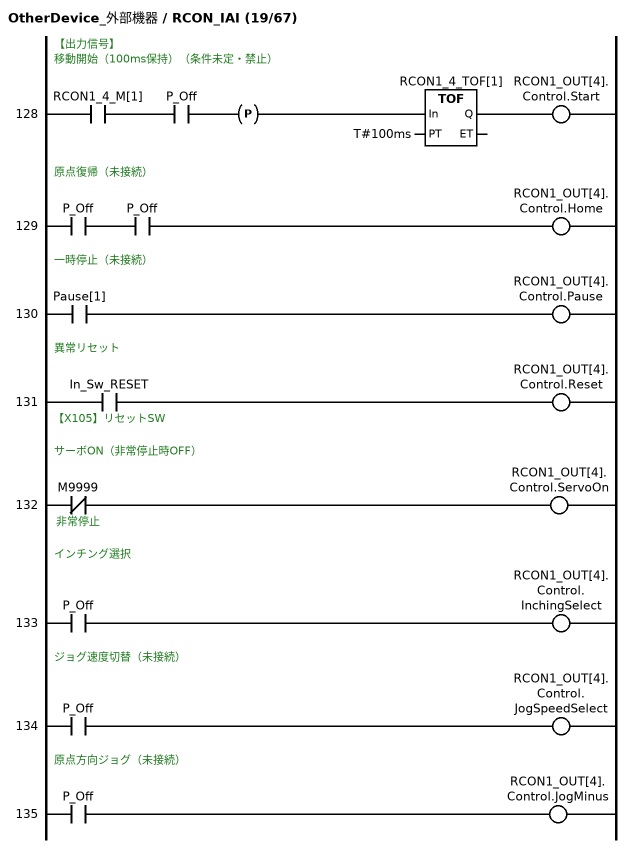
(* [picture p96: OtherDevice_外部機器 / RCON_IAI, rungs 128-135] *)
(* Rung 128: 【出力信号】 / 移動開始（100ms保持）（条件未定・禁止） *)
_e13(CLK := RCON1_4_M[1] AND P_Off);
RCON1_4_TOF[1](In := _e13.Q, PT := T#100ms);
RCON1_OUT[4].Control.Start := RCON1_4_TOF[1].Q;
(* Rung 129: 原点復帰（未接続） *)
RCON1_OUT[4].Control.Home := P_Off AND P_Off;
(* Rung 130: 一時停止（未接続） *)
RCON1_OUT[4].Control.Pause := Pause[1];
(* Rung 131: 異常リセット *)
RCON1_OUT[4].Control.Reset := In_Sw_RESET;
(* Rung 132: サーボON（非常停止時OFF） *)
RCON1_OUT[4].Control.ServoOn := NOT M9999;
(* Rung 133: インチング選択 *)
RCON1_OUT[4].Control.InchingSelect := P_Off;
(* Rung 134: ジョグ速度切替（未接続） *)
RCON1_OUT[4].Control.JogSpeedSelect := P_Off;
(* Rung 135: 原点方向ジョグ（未接続） *)
RCON1_OUT[4].Control.JogMinus := P_Off;

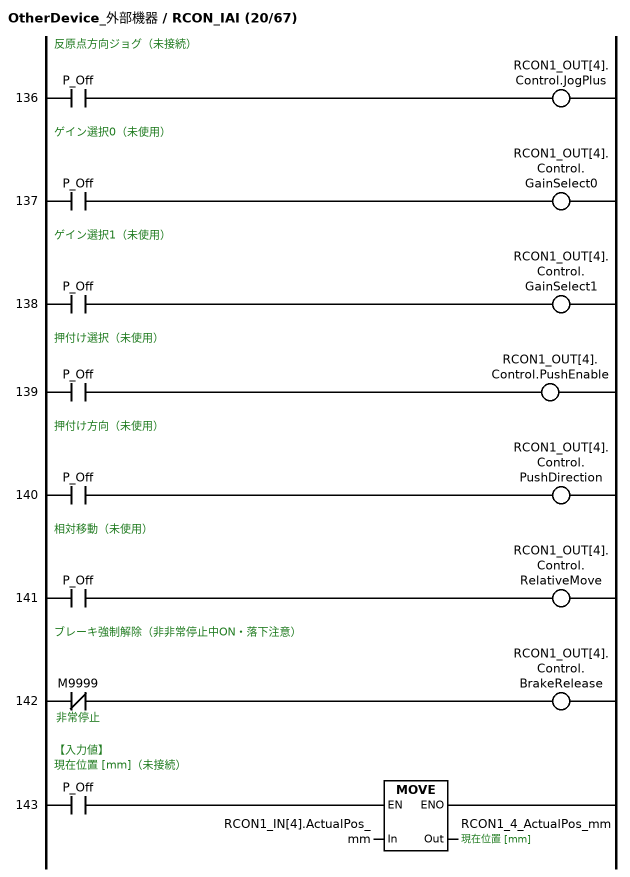
(* Rung 136: 反原点方向ジョグ（未接続） *)
RCON1_OUT[4].Control.JogPlus := P_Off;
(* Rung 137: ゲイン選択0（未使用） *)
RCON1_OUT[4].Control.GainSelect0 := P_Off;
(* Rung 138: ゲイン選択1（未使用） *)
RCON1_OUT[4].Control.GainSelect1 := P_Off;
(* Rung 139: 押付け選択（未使用） *)
RCON1_OUT[4].Control.PushEnable := P_Off;
(* Rung 140: 押付け方向（未使用） *)
RCON1_OUT[4].Control.PushDirection := P_Off;
(* Rung 141: 相対移動（未使用） *)
RCON1_OUT[4].Control.RelativeMove := P_Off;
(* Rung 142: ブレーキ強制解除（非非常停止中ON・落下注意） *)
RCON1_OUT[4].Control.BrakeRelease := NOT M9999;
(* Rung 143: 【入力値】 / 現在位置 [mm]（未接続） *)
IF P_Off THEN RCON1_4_ActualPos_mm := RCON1_IN[4].ActualPos_mm; END_IF;

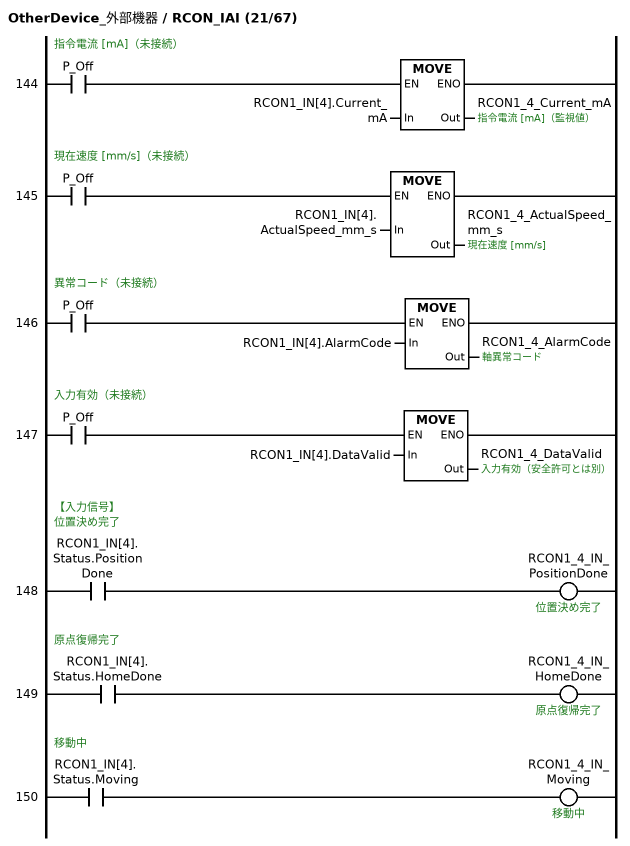
(* Rung 144: 指令電流 [mA]（未接続） *)
IF P_Off THEN RCON1_4_Current_mA := RCON1_IN[4].Current_mA; END_IF;
(* Rung 145: 現在速度 [mm/s]（未接続） *)
IF P_Off THEN RCON1_4_ActualSpeed_mm_s := RCON1_IN[4].ActualSpeed_mm_s; END_IF;
(* Rung 146: 異常コード（未接続） *)
IF P_Off THEN RCON1_4_AlarmCode := RCON1_IN[4].AlarmCode; END_IF;
(* Rung 147: 入力有効（未接続） *)
IF P_Off THEN RCON1_4_DataValid := RCON1_IN[4].DataValid; END_IF;
(* Rung 148: 【入力信号】 / 位置決め完了 *)
RCON1_4_IN_PositionDone := RCON1_IN[4].Status.PositionDone;
(* Rung 149: 原点復帰完了 *)
RCON1_4_IN_HomeDone := RCON1_IN[4].Status.HomeDone;
(* Rung 150: 移動中 *)
RCON1_4_IN_Moving := RCON1_IN[4].Status.Moving;

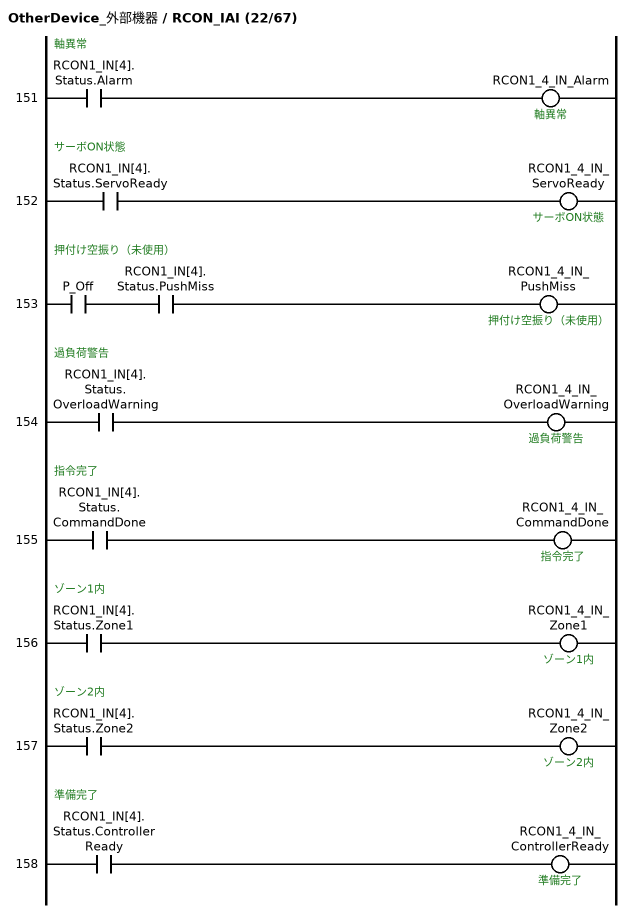
(* Rung 151: 軸異常 *)
RCON1_4_IN_Alarm := RCON1_IN[4].Status.Alarm;
(* Rung 152: サーボON状態 *)
RCON1_4_IN_ServoReady := RCON1_IN[4].Status.ServoReady;
(* Rung 153: 押付け空振り（未使用） *)
RCON1_4_IN_PushMiss := P_Off AND RCON1_IN[4].Status.PushMiss;
(* Rung 154: 過負荷警告 *)
RCON1_4_IN_OverloadWarning := RCON1_IN[4].Status.OverloadWarning;
(* Rung 155: 指令完了 *)
RCON1_4_IN_CommandDone := RCON1_IN[4].Status.CommandDone;
(* Rung 156: ゾーン1内 *)
RCON1_4_IN_Zone1 := RCON1_IN[4].Status.Zone1;
(* Rung 157: ゾーン2内 *)
RCON1_4_IN_Zone2 := RCON1_IN[4].Status.Zone2;
(* Rung 158: 準備完了 *)
RCON1_4_IN_ControllerReady := RCON1_IN[4].Status.ControllerReady;

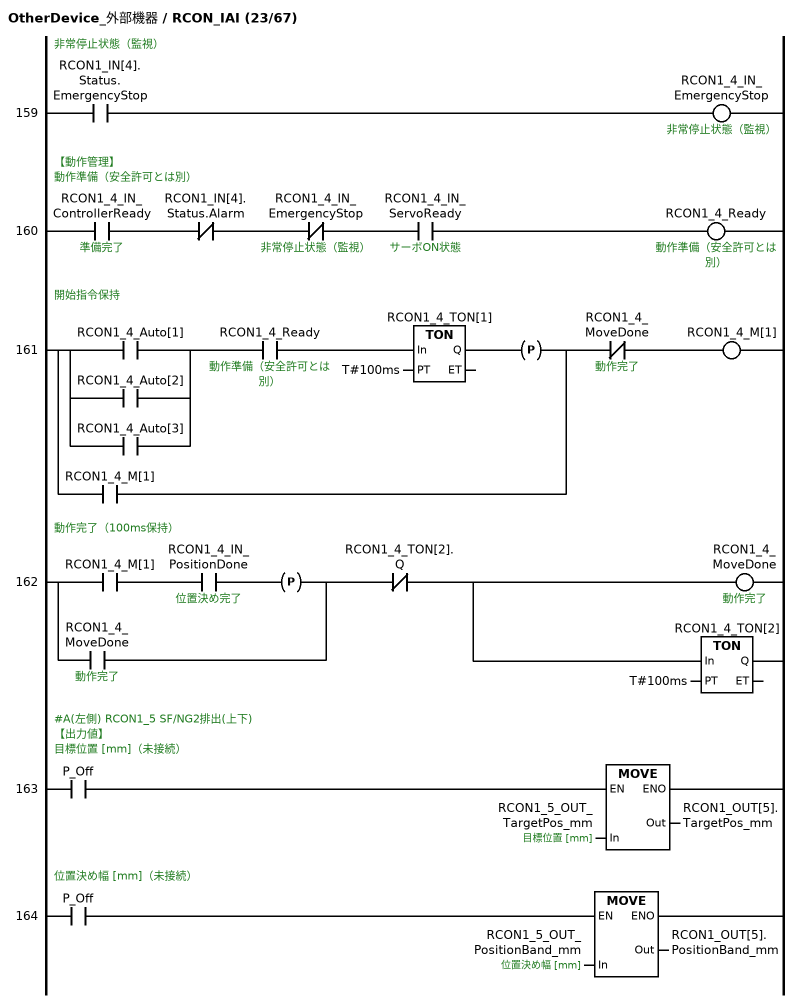
(* Rung 159: 非常停止状態（監視） *)
RCON1_4_IN_EmergencyStop := RCON1_IN[4].Status.EmergencyStop;
(* Rung 160: 【動作管理】 / 動作準備（安全許可とは別） *)
RCON1_4_Ready := RCON1_4_IN_ControllerReady AND NOT RCON1_IN[4].Status.Alarm AND NOT RCON1_4_IN_EmergencyStop AND RCON1_4_IN_ServoReady;
(* Rung 161: 開始指令保持 *)
RCON1_4_TON[1](In := (RCON1_4_Auto[1] OR RCON1_4_Auto[2] OR RCON1_4_Auto[3]) AND RCON1_4_Ready, PT := T#100ms);
_e14(CLK := RCON1_4_TON[1].Q);
RCON1_4_M[1] := (_e14.Q OR RCON1_4_M[1]) AND NOT RCON1_4_MoveDone;
(* Rung 162: 動作完了（100ms保持） *)
_e15(CLK := RCON1_4_M[1] AND RCON1_4_IN_PositionDone);
_p16 := (_e15.Q OR RCON1_4_MoveDone) AND NOT RCON1_4_TON[2].Q;
RCON1_4_MoveDone := _p16;
RCON1_4_TON[2](In := _p16, PT := T#100ms);
(* Rung 163: #A(左側) RCON1_5 SF/NG2排出(上下) / 【出力値】 / 目標位置 [mm]（未接続） *)
IF P_Off THEN RCON1_OUT[5].TargetPos_mm := RCON1_5_OUT_TargetPos_mm; END_IF;
(* Rung 164: 位置決め幅 [mm]（未接続） *)
IF P_Off THEN RCON1_OUT[5].PositionBand_mm := RCON1_5_OUT_PositionBand_mm; END_IF;

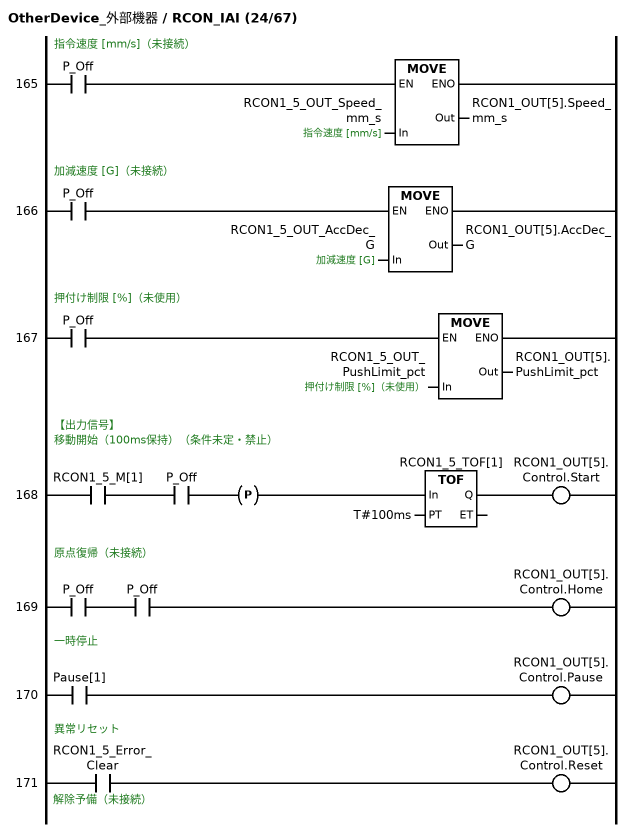
(* Rung 165: 指令速度 [mm/s]（未接続） *)
IF P_Off THEN RCON1_OUT[5].Speed_mm_s := RCON1_5_OUT_Speed_mm_s; END_IF;
(* Rung 166: 加減速度 [G]（未接続） *)
IF P_Off THEN RCON1_OUT[5].AccDec_G := RCON1_5_OUT_AccDec_G; END_IF;
(* Rung 167: 押付け制限 [%]（未使用） *)
IF P_Off THEN RCON1_OUT[5].PushLimit_pct := RCON1_5_OUT_PushLimit_pct; END_IF;
(* Rung 168: 【出力信号】 / 移動開始（100ms保持）（条件未定・禁止） *)
_e17(CLK := RCON1_5_M[1] AND P_Off);
RCON1_5_TOF[1](In := _e17.Q, PT := T#100ms);
RCON1_OUT[5].Control.Start := RCON1_5_TOF[1].Q;
(* Rung 169: 原点復帰（未接続） *)
RCON1_OUT[5].Control.Home := P_Off AND P_Off;
(* Rung 170: 一時停止 *)
RCON1_OUT[5].Control.Pause := Pause[1];
(* Rung 171: 異常リセット *)
RCON1_OUT[5].Control.Reset := RCON1_5_Error_Clear;

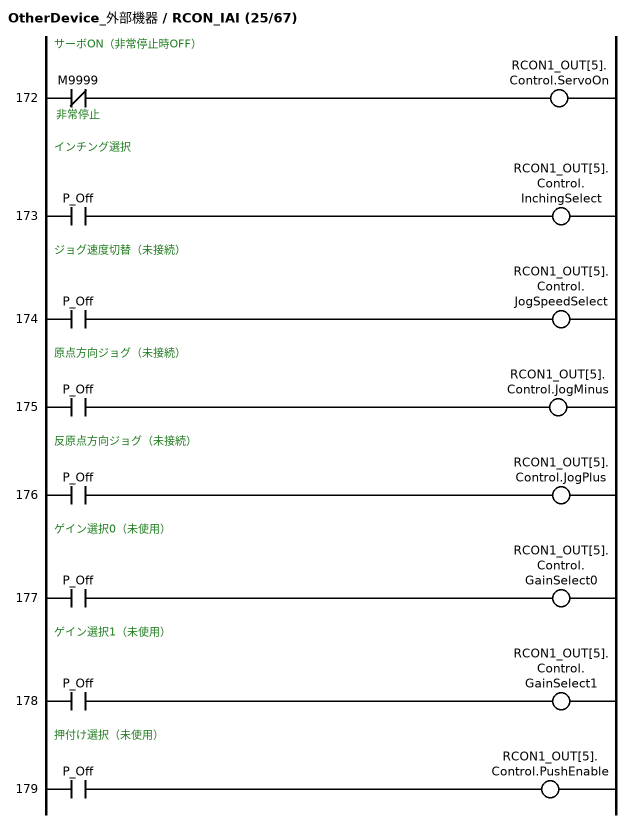
(* Rung 172: サーボON（非常停止時OFF） *)
RCON1_OUT[5].Control.ServoOn := NOT M9999;
(* Rung 173: インチング選択 *)
RCON1_OUT[5].Control.InchingSelect := P_Off;
(* Rung 174: ジョグ速度切替（未接続） *)
RCON1_OUT[5].Control.JogSpeedSelect := P_Off;
(* Rung 175: 原点方向ジョグ（未接続） *)
RCON1_OUT[5].Control.JogMinus := P_Off;
(* Rung 176: 反原点方向ジョグ（未接続） *)
RCON1_OUT[5].Control.JogPlus := P_Off;
(* Rung 177: ゲイン選択0（未使用） *)
RCON1_OUT[5].Control.GainSelect0 := P_Off;
(* Rung 178: ゲイン選択1（未使用） *)
RCON1_OUT[5].Control.GainSelect1 := P_Off;
(* Rung 179: 押付け選択（未使用） *)
RCON1_OUT[5].Control.PushEnable := P_Off;

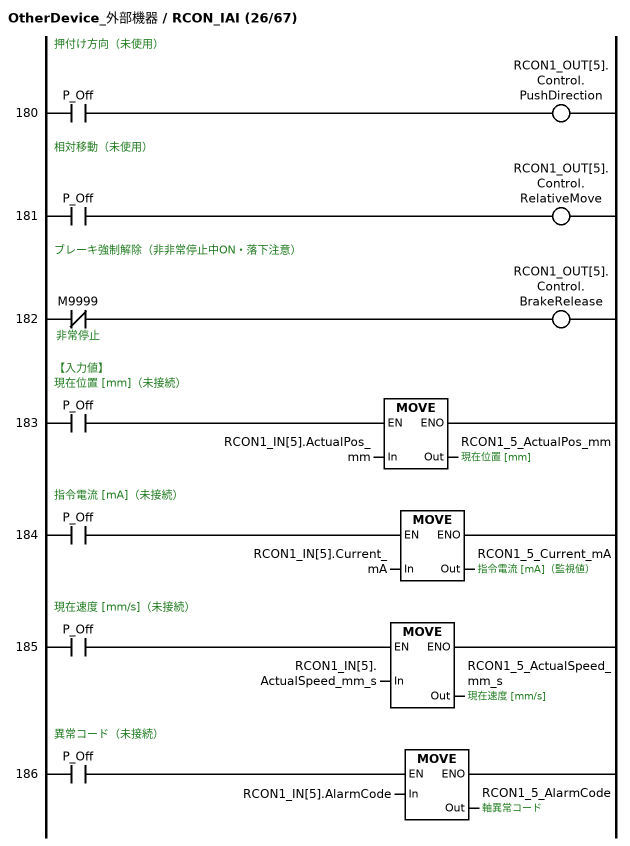
(* Rung 180: 押付け方向（未使用） *)
RCON1_OUT[5].Control.PushDirection := P_Off;
(* Rung 181: 相対移動（未使用） *)
RCON1_OUT[5].Control.RelativeMove := P_Off;
(* Rung 182: ブレーキ強制解除（非非常停止中ON・落下注意） *)
RCON1_OUT[5].Control.BrakeRelease := NOT M9999;
(* Rung 183: 【入力値】 / 現在位置 [mm]（未接続） *)
IF P_Off THEN RCON1_5_ActualPos_mm := RCON1_IN[5].ActualPos_mm; END_IF;
(* Rung 184: 指令電流 [mA]（未接続） *)
IF P_Off THEN RCON1_5_Current_mA := RCON1_IN[5].Current_mA; END_IF;
(* Rung 185: 現在速度 [mm/s]（未接続） *)
IF P_Off THEN RCON1_5_ActualSpeed_mm_s := RCON1_IN[5].ActualSpeed_mm_s; END_IF;
(* Rung 186: 異常コード（未接続） *)
IF P_Off THEN RCON1_5_AlarmCode := RCON1_IN[5].AlarmCode; END_IF;

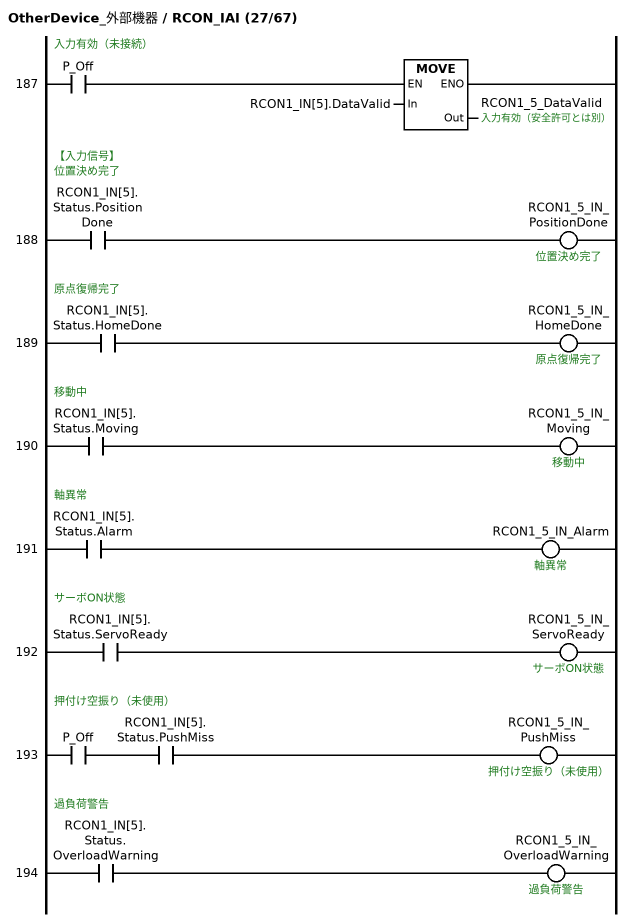
(* Rung 187: 入力有効（未接続） *)
IF P_Off THEN RCON1_5_DataValid := RCON1_IN[5].DataValid; END_IF;
(* Rung 188: 【入力信号】 / 位置決め完了 *)
RCON1_5_IN_PositionDone := RCON1_IN[5].Status.PositionDone;
(* Rung 189: 原点復帰完了 *)
RCON1_5_IN_HomeDone := RCON1_IN[5].Status.HomeDone;
(* Rung 190: 移動中 *)
RCON1_5_IN_Moving := RCON1_IN[5].Status.Moving;
(* Rung 191: 軸異常 *)
RCON1_5_IN_Alarm := RCON1_IN[5].Status.Alarm;
(* Rung 192: サーボON状態 *)
RCON1_5_IN_ServoReady := RCON1_IN[5].Status.ServoReady;
(* Rung 193: 押付け空振り（未使用） *)
RCON1_5_IN_PushMiss := P_Off AND RCON1_IN[5].Status.PushMiss;
(* Rung 194: 過負荷警告 *)
RCON1_5_IN_OverloadWarning := RCON1_IN[5].Status.OverloadWarning;

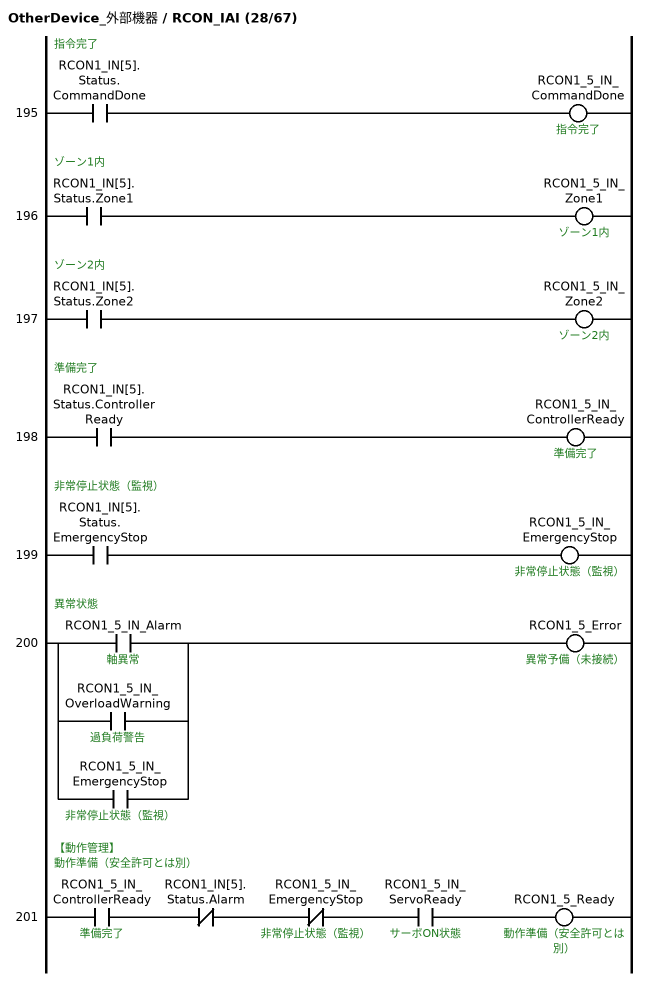
(* Rung 195: 指令完了 *)
RCON1_5_IN_CommandDone := RCON1_IN[5].Status.CommandDone;
(* Rung 196: ゾーン1内 *)
RCON1_5_IN_Zone1 := RCON1_IN[5].Status.Zone1;
(* Rung 197: ゾーン2内 *)
RCON1_5_IN_Zone2 := RCON1_IN[5].Status.Zone2;
(* Rung 198: 準備完了 *)
RCON1_5_IN_ControllerReady := RCON1_IN[5].Status.ControllerReady;
(* Rung 199: 非常停止状態（監視） *)
RCON1_5_IN_EmergencyStop := RCON1_IN[5].Status.EmergencyStop;
(* Rung 200: 異常状態 *)
RCON1_5_Error := RCON1_5_IN_Alarm OR RCON1_5_IN_OverloadWarning OR RCON1_5_IN_EmergencyStop;
(* Rung 201: 【動作管理】 / 動作準備（安全許可とは別） *)
RCON1_5_Ready := RCON1_5_IN_ControllerReady AND NOT RCON1_IN[5].Status.Alarm AND NOT RCON1_5_IN_EmergencyStop AND RCON1_5_IN_ServoReady;

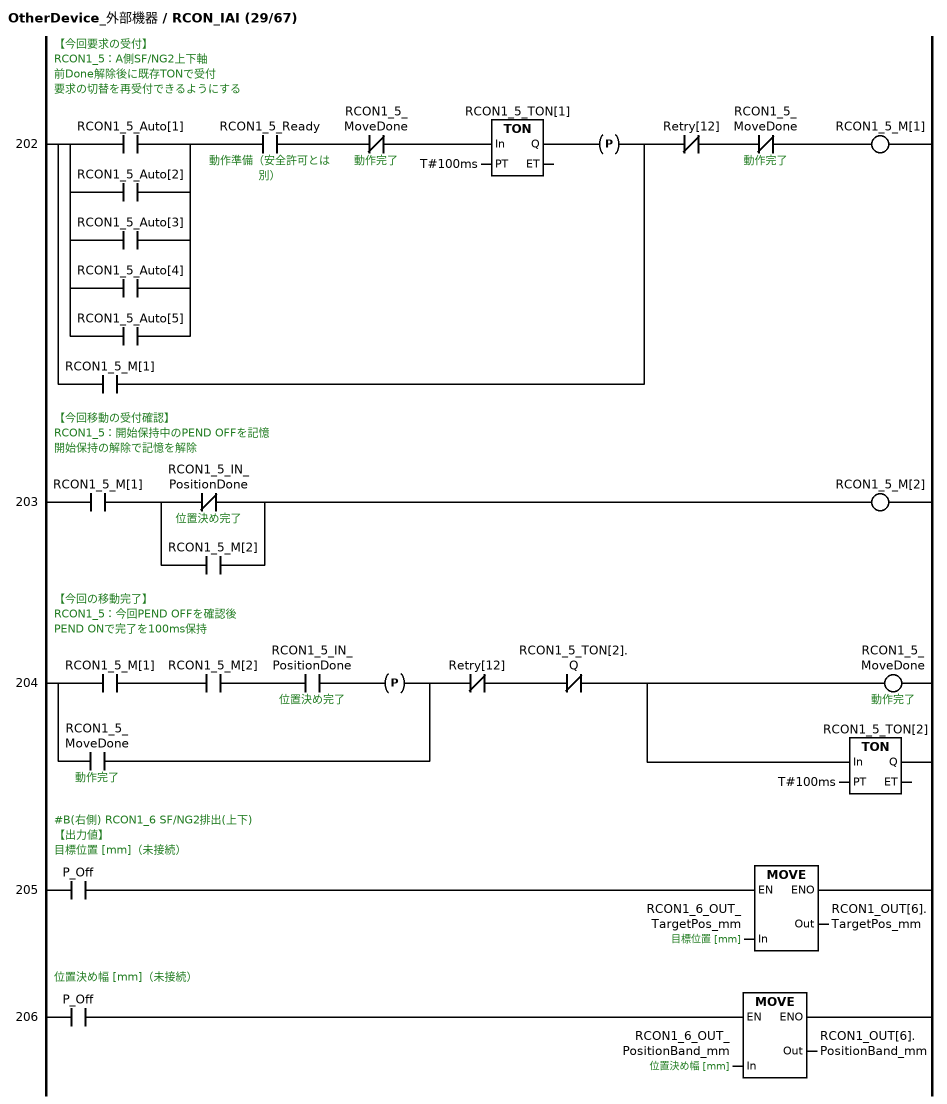
(* Rung 202: 【今回要求の受付】 / RCON1_5：A側SF/NG2上下軸 / 前Done解除後に既存TONで受付 / 要求の切替を再受付できるようにする *)
RCON1_5_TON[1](In := (RCON1_5_Auto[1] OR RCON1_5_Auto[2] OR RCON1_5_Auto[3] OR RCON1_5_Auto[4] OR RCON1_5_Auto[5]) AND RCON1_5_Ready AND NOT RCON1_5_MoveDone, PT := T#100ms);
_e18(CLK := RCON1_5_TON[1].Q);
RCON1_5_M[1] := (_e18.Q OR RCON1_5_M[1]) AND NOT Retry[12] AND NOT RCON1_5_MoveDone;
(* Rung 203: 【今回移動の受付確認】 / RCON1_5：開始保持中のPEND OFFを記憶 / 開始保持の解除で記憶を解除 *)
RCON1_5_M[2] := RCON1_5_M[1] AND (NOT RCON1_5_IN_PositionDone OR RCON1_5_M[2]);
(* Rung 204: 【今回の移動完了】 / RCON1_5：今回PEND OFFを確認後 / PEND ONで完了を100ms保持 *)
_e19(CLK := RCON1_5_M[1] AND RCON1_5_M[2] AND RCON1_5_IN_PositionDone);
_p20 := (_e19.Q OR RCON1_5_MoveDone) AND NOT Retry[12] AND NOT RCON1_5_TON[2].Q;
RCON1_5_MoveDone := _p20;
RCON1_5_TON[2](In := _p20, PT := T#100ms);
(* Rung 205: #B(右側) RCON1_6 SF/NG2排出(上下) / 【出力値】 / 目標位置 [mm]（未接続） *)
IF P_Off THEN RCON1_OUT[6].TargetPos_mm := RCON1_6_OUT_TargetPos_mm; END_IF;
(* Rung 206: 位置決め幅 [mm]（未接続） *)
IF P_Off THEN RCON1_OUT[6].PositionBand_mm := RCON1_6_OUT_PositionBand_mm; END_IF;

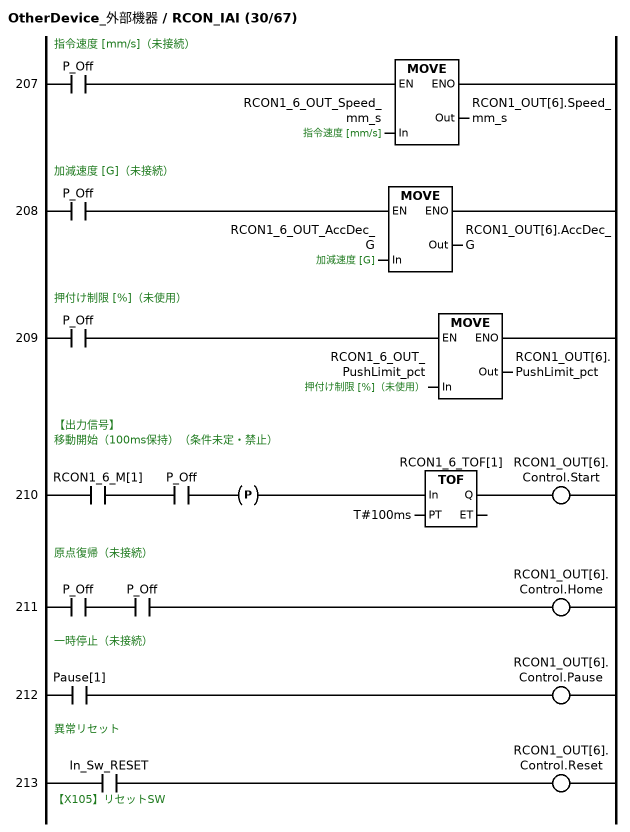
(* Rung 207: 指令速度 [mm/s]（未接続） *)
IF P_Off THEN RCON1_OUT[6].Speed_mm_s := RCON1_6_OUT_Speed_mm_s; END_IF;
(* Rung 208: 加減速度 [G]（未接続） *)
IF P_Off THEN RCON1_OUT[6].AccDec_G := RCON1_6_OUT_AccDec_G; END_IF;
(* Rung 209: 押付け制限 [%]（未使用） *)
IF P_Off THEN RCON1_OUT[6].PushLimit_pct := RCON1_6_OUT_PushLimit_pct; END_IF;
(* Rung 210: 【出力信号】 / 移動開始（100ms保持）（条件未定・禁止） *)
_e21(CLK := RCON1_6_M[1] AND P_Off);
RCON1_6_TOF[1](In := _e21.Q, PT := T#100ms);
RCON1_OUT[6].Control.Start := RCON1_6_TOF[1].Q;
(* Rung 211: 原点復帰（未接続） *)
RCON1_OUT[6].Control.Home := P_Off AND P_Off;
(* Rung 212: 一時停止（未接続） *)
RCON1_OUT[6].Control.Pause := Pause[1];
(* Rung 213: 異常リセット *)
RCON1_OUT[6].Control.Reset := In_Sw_RESET;

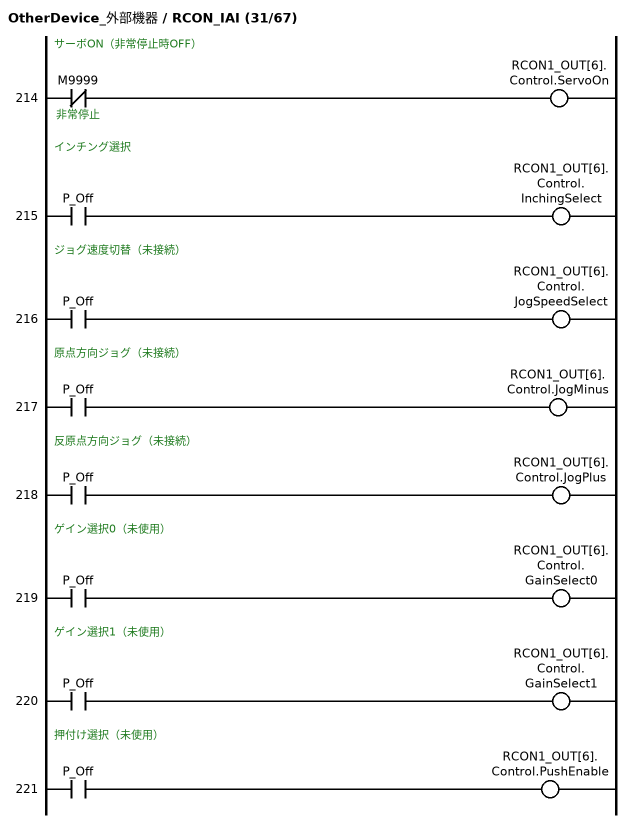
(* Rung 214: サーボON（非常停止時OFF） *)
RCON1_OUT[6].Control.ServoOn := NOT M9999;
(* Rung 215: インチング選択 *)
RCON1_OUT[6].Control.InchingSelect := P_Off;
(* Rung 216: ジョグ速度切替（未接続） *)
RCON1_OUT[6].Control.JogSpeedSelect := P_Off;
(* Rung 217: 原点方向ジョグ（未接続） *)
RCON1_OUT[6].Control.JogMinus := P_Off;
(* Rung 218: 反原点方向ジョグ（未接続） *)
RCON1_OUT[6].Control.JogPlus := P_Off;
(* Rung 219: ゲイン選択0（未使用） *)
RCON1_OUT[6].Control.GainSelect0 := P_Off;
(* Rung 220: ゲイン選択1（未使用） *)
RCON1_OUT[6].Control.GainSelect1 := P_Off;
(* Rung 221: 押付け選択（未使用） *)
RCON1_OUT[6].Control.PushEnable := P_Off;

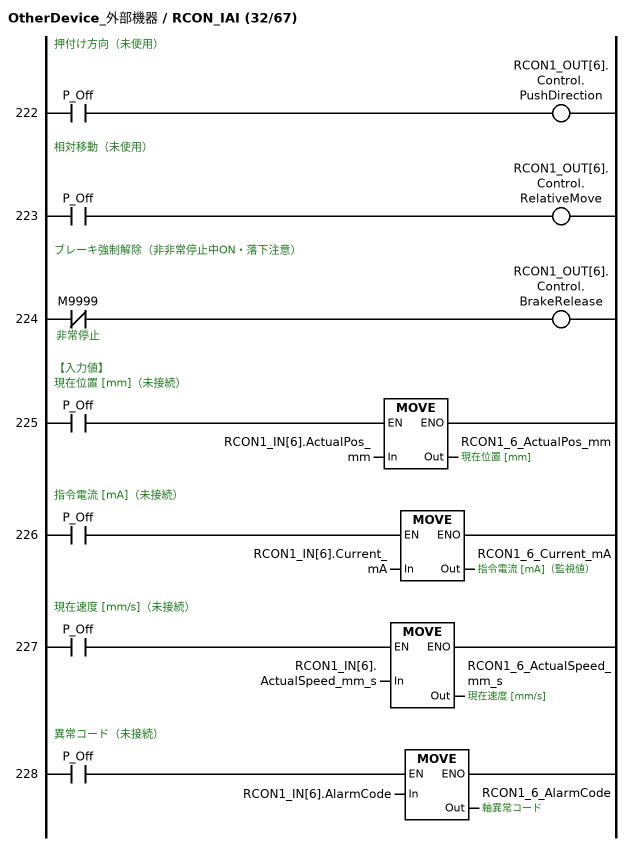
(* Rung 222: 押付け方向（未使用） *)
RCON1_OUT[6].Control.PushDirection := P_Off;
(* Rung 223: 相対移動（未使用） *)
RCON1_OUT[6].Control.RelativeMove := P_Off;
(* Rung 224: ブレーキ強制解除（非非常停止中ON・落下注意） *)
RCON1_OUT[6].Control.BrakeRelease := NOT M9999;
(* Rung 225: 【入力値】 / 現在位置 [mm]（未接続） *)
IF P_Off THEN RCON1_6_ActualPos_mm := RCON1_IN[6].ActualPos_mm; END_IF;
(* Rung 226: 指令電流 [mA]（未接続） *)
IF P_Off THEN RCON1_6_Current_mA := RCON1_IN[6].Current_mA; END_IF;
(* Rung 227: 現在速度 [mm/s]（未接続） *)
IF P_Off THEN RCON1_6_ActualSpeed_mm_s := RCON1_IN[6].ActualSpeed_mm_s; END_IF;
(* Rung 228: 異常コード（未接続） *)
IF P_Off THEN RCON1_6_AlarmCode := RCON1_IN[6].AlarmCode; END_IF;

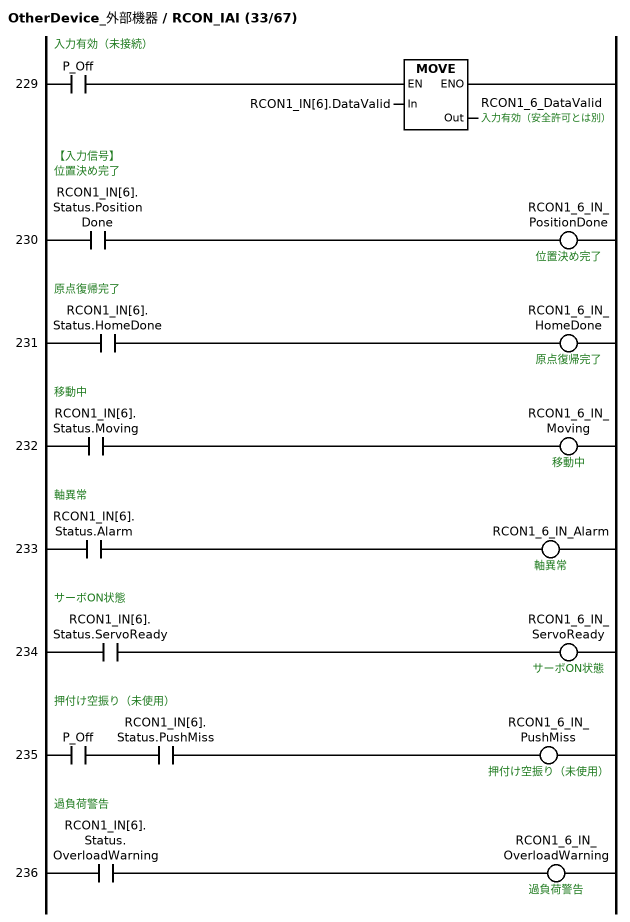
(* Rung 229: 入力有効（未接続） *)
IF P_Off THEN RCON1_6_DataValid := RCON1_IN[6].DataValid; END_IF;
(* Rung 230: 【入力信号】 / 位置決め完了 *)
RCON1_6_IN_PositionDone := RCON1_IN[6].Status.PositionDone;
(* Rung 231: 原点復帰完了 *)
RCON1_6_IN_HomeDone := RCON1_IN[6].Status.HomeDone;
(* Rung 232: 移動中 *)
RCON1_6_IN_Moving := RCON1_IN[6].Status.Moving;
(* Rung 233: 軸異常 *)
RCON1_6_IN_Alarm := RCON1_IN[6].Status.Alarm;
(* Rung 234: サーボON状態 *)
RCON1_6_IN_ServoReady := RCON1_IN[6].Status.ServoReady;
(* Rung 235: 押付け空振り（未使用） *)
RCON1_6_IN_PushMiss := P_Off AND RCON1_IN[6].Status.PushMiss;
(* Rung 236: 過負荷警告 *)
RCON1_6_IN_OverloadWarning := RCON1_IN[6].Status.OverloadWarning;

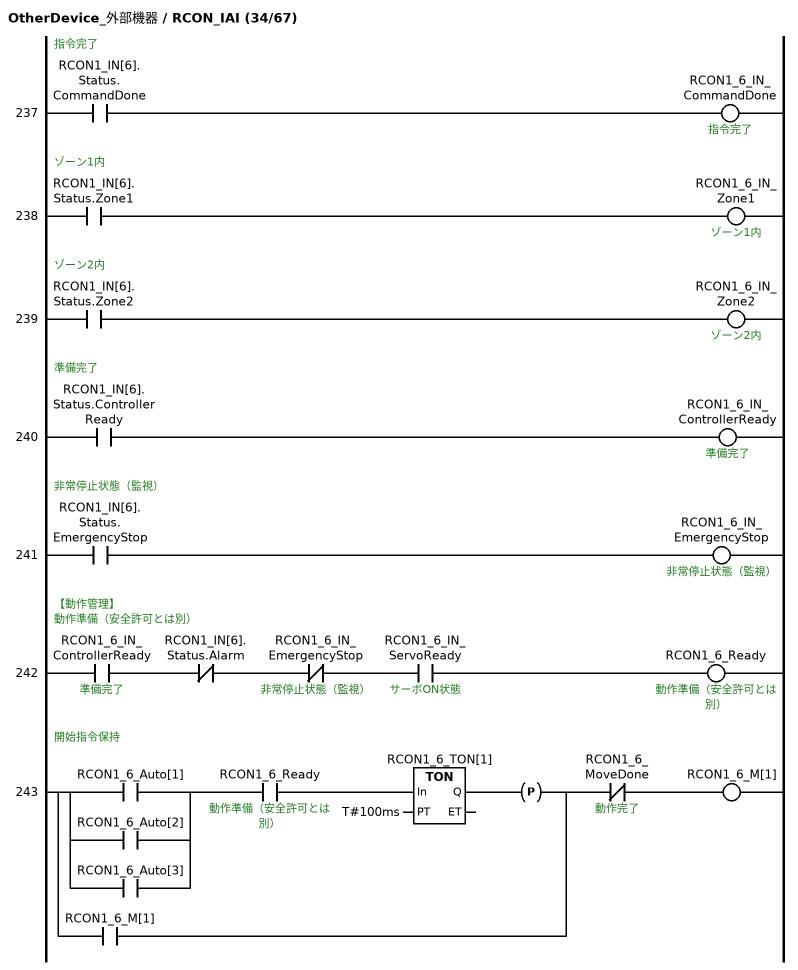
(* Rung 237: 指令完了 *)
RCON1_6_IN_CommandDone := RCON1_IN[6].Status.CommandDone;
(* Rung 238: ゾーン1内 *)
RCON1_6_IN_Zone1 := RCON1_IN[6].Status.Zone1;
(* Rung 239: ゾーン2内 *)
RCON1_6_IN_Zone2 := RCON1_IN[6].Status.Zone2;
(* Rung 240: 準備完了 *)
RCON1_6_IN_ControllerReady := RCON1_IN[6].Status.ControllerReady;
(* Rung 241: 非常停止状態（監視） *)
RCON1_6_IN_EmergencyStop := RCON1_IN[6].Status.EmergencyStop;
(* Rung 242: 【動作管理】 / 動作準備（安全許可とは別） *)
RCON1_6_Ready := RCON1_6_IN_ControllerReady AND NOT RCON1_IN[6].Status.Alarm AND NOT RCON1_6_IN_EmergencyStop AND RCON1_6_IN_ServoReady;
(* Rung 243: 開始指令保持 *)
RCON1_6_TON[1](In := (RCON1_6_Auto[1] OR RCON1_6_Auto[2] OR RCON1_6_Auto[3]) AND RCON1_6_Ready, PT := T#100ms);
_e22(CLK := RCON1_6_TON[1].Q);
RCON1_6_M[1] := (_e22.Q OR RCON1_6_M[1]) AND NOT RCON1_6_MoveDone;

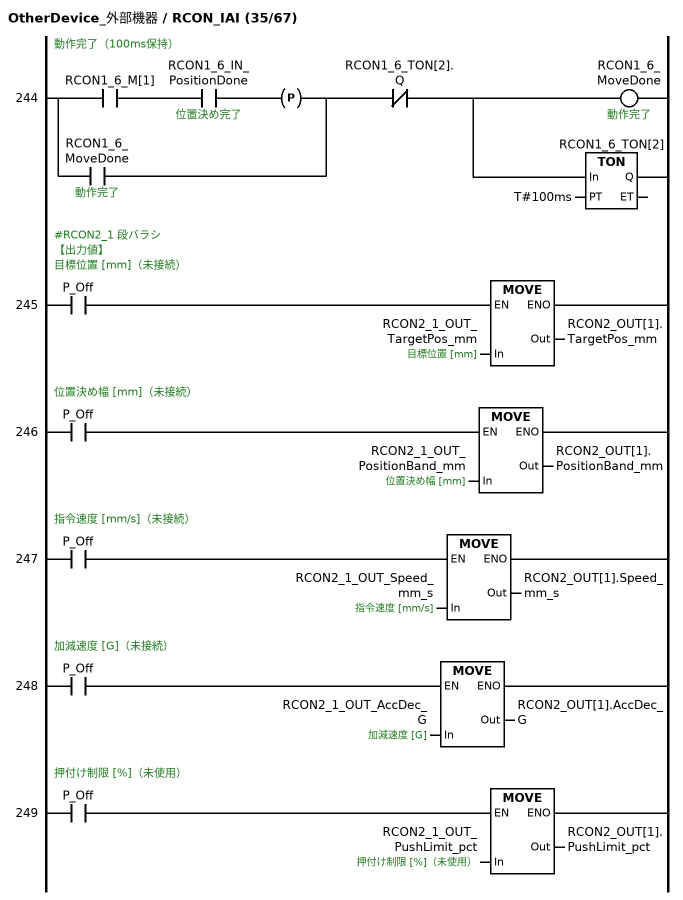
(* Rung 244: 動作完了（100ms保持） *)
_e23(CLK := RCON1_6_M[1] AND RCON1_6_IN_PositionDone);
_p24 := (_e23.Q OR RCON1_6_MoveDone) AND NOT RCON1_6_TON[2].Q;
RCON1_6_MoveDone := _p24;
RCON1_6_TON[2](In := _p24, PT := T#100ms);
(* Rung 245: #RCON2_1 段バラシ / 【出力値】 / 目標位置 [mm]（未接続） *)
IF P_Off THEN RCON2_OUT[1].TargetPos_mm := RCON2_1_OUT_TargetPos_mm; END_IF;
(* Rung 246: 位置決め幅 [mm]（未接続） *)
IF P_Off THEN RCON2_OUT[1].PositionBand_mm := RCON2_1_OUT_PositionBand_mm; END_IF;
(* Rung 247: 指令速度 [mm/s]（未接続） *)
IF P_Off THEN RCON2_OUT[1].Speed_mm_s := RCON2_1_OUT_Speed_mm_s; END_IF;
(* Rung 248: 加減速度 [G]（未接続） *)
IF P_Off THEN RCON2_OUT[1].AccDec_G := RCON2_1_OUT_AccDec_G; END_IF;
(* Rung 249: 押付け制限 [%]（未使用） *)
IF P_Off THEN RCON2_OUT[1].PushLimit_pct := RCON2_1_OUT_PushLimit_pct; END_IF;

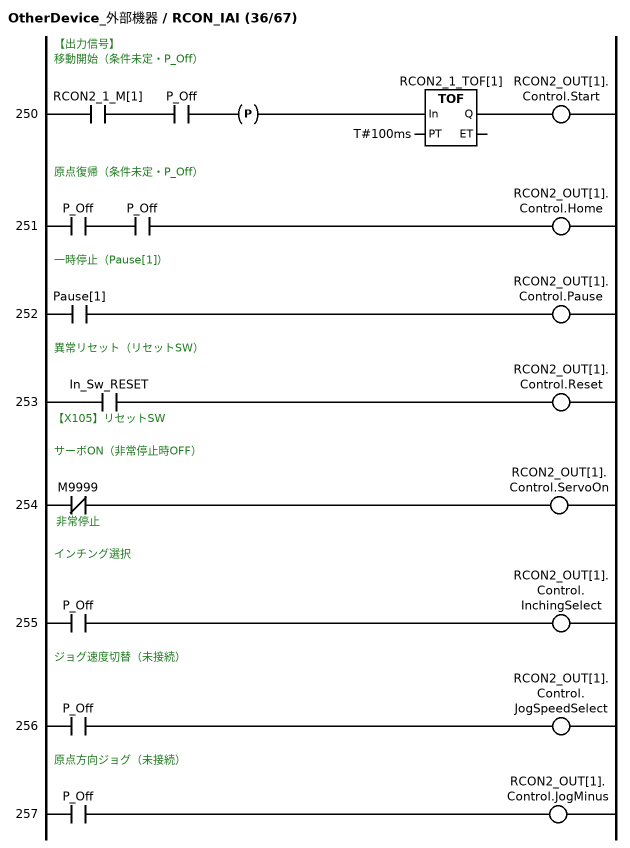
(* Rung 250: 【出力信号】 / 移動開始（条件未定・P_Off） *)
_e25(CLK := RCON2_1_M[1] AND P_Off);
RCON2_1_TOF[1](In := _e25.Q, PT := T#100ms);
RCON2_OUT[1].Control.Start := RCON2_1_TOF[1].Q;
(* Rung 251: 原点復帰（条件未定・P_Off） *)
RCON2_OUT[1].Control.Home := P_Off AND P_Off;
(* Rung 252: 一時停止（Pause[1]） *)
RCON2_OUT[1].Control.Pause := Pause[1];
(* Rung 253: 異常リセット（リセットSW） *)
RCON2_OUT[1].Control.Reset := In_Sw_RESET;
(* Rung 254: サーボON（非常停止時OFF） *)
RCON2_OUT[1].Control.ServoOn := NOT M9999;
(* Rung 255: インチング選択 *)
RCON2_OUT[1].Control.InchingSelect := P_Off;
(* Rung 256: ジョグ速度切替（未接続） *)
RCON2_OUT[1].Control.JogSpeedSelect := P_Off;
(* Rung 257: 原点方向ジョグ（未接続） *)
RCON2_OUT[1].Control.JogMinus := P_Off;

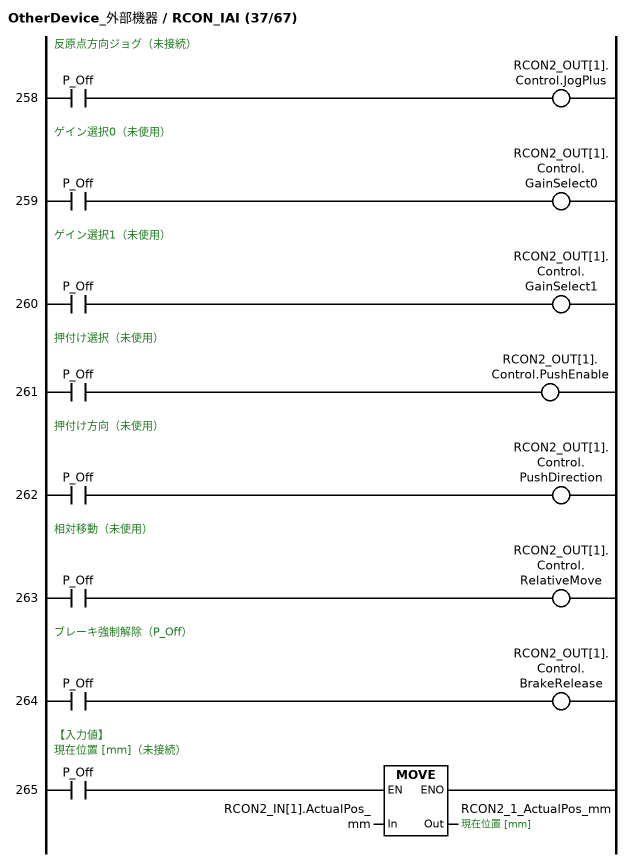
(* Rung 258: 反原点方向ジョグ（未接続） *)
RCON2_OUT[1].Control.JogPlus := P_Off;
(* Rung 259: ゲイン選択0（未使用） *)
RCON2_OUT[1].Control.GainSelect0 := P_Off;
(* Rung 260: ゲイン選択1（未使用） *)
RCON2_OUT[1].Control.GainSelect1 := P_Off;
(* Rung 261: 押付け選択（未使用） *)
RCON2_OUT[1].Control.PushEnable := P_Off;
(* Rung 262: 押付け方向（未使用） *)
RCON2_OUT[1].Control.PushDirection := P_Off;
(* Rung 263: 相対移動（未使用） *)
RCON2_OUT[1].Control.RelativeMove := P_Off;
(* Rung 264: ブレーキ強制解除（P_Off） *)
RCON2_OUT[1].Control.BrakeRelease := P_Off;
(* Rung 265: 【入力値】 / 現在位置 [mm]（未接続） *)
IF P_Off THEN RCON2_1_ActualPos_mm := RCON2_IN[1].ActualPos_mm; END_IF;

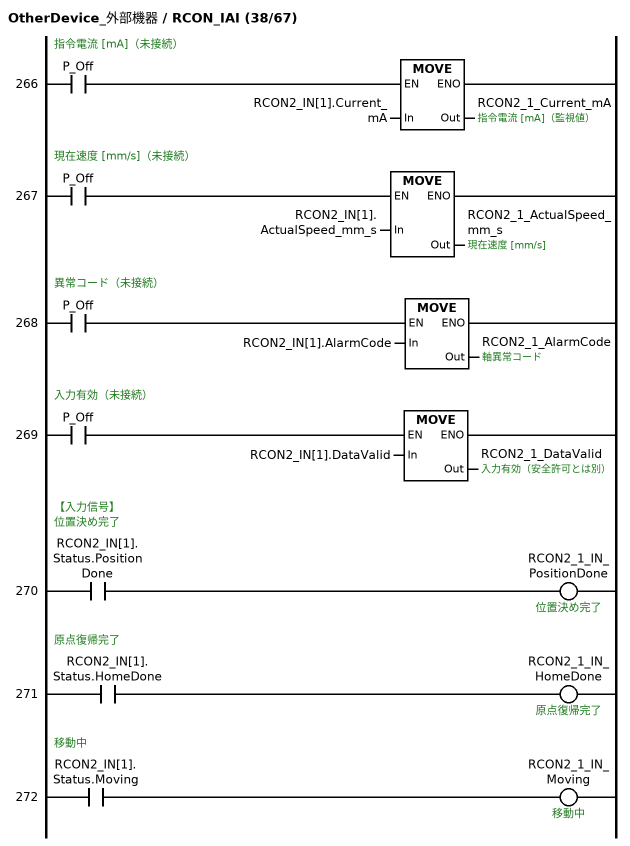
(* Rung 266: 指令電流 [mA]（未接続） *)
IF P_Off THEN RCON2_1_Current_mA := RCON2_IN[1].Current_mA; END_IF;
(* Rung 267: 現在速度 [mm/s]（未接続） *)
IF P_Off THEN RCON2_1_ActualSpeed_mm_s := RCON2_IN[1].ActualSpeed_mm_s; END_IF;
(* Rung 268: 異常コード（未接続） *)
IF P_Off THEN RCON2_1_AlarmCode := RCON2_IN[1].AlarmCode; END_IF;
(* Rung 269: 入力有効（未接続） *)
IF P_Off THEN RCON2_1_DataValid := RCON2_IN[1].DataValid; END_IF;
(* Rung 270: 【入力信号】 / 位置決め完了 *)
RCON2_1_IN_PositionDone := RCON2_IN[1].Status.PositionDone;
(* Rung 271: 原点復帰完了 *)
RCON2_1_IN_HomeDone := RCON2_IN[1].Status.HomeDone;
(* Rung 272: 移動中 *)
RCON2_1_IN_Moving := RCON2_IN[1].Status.Moving;

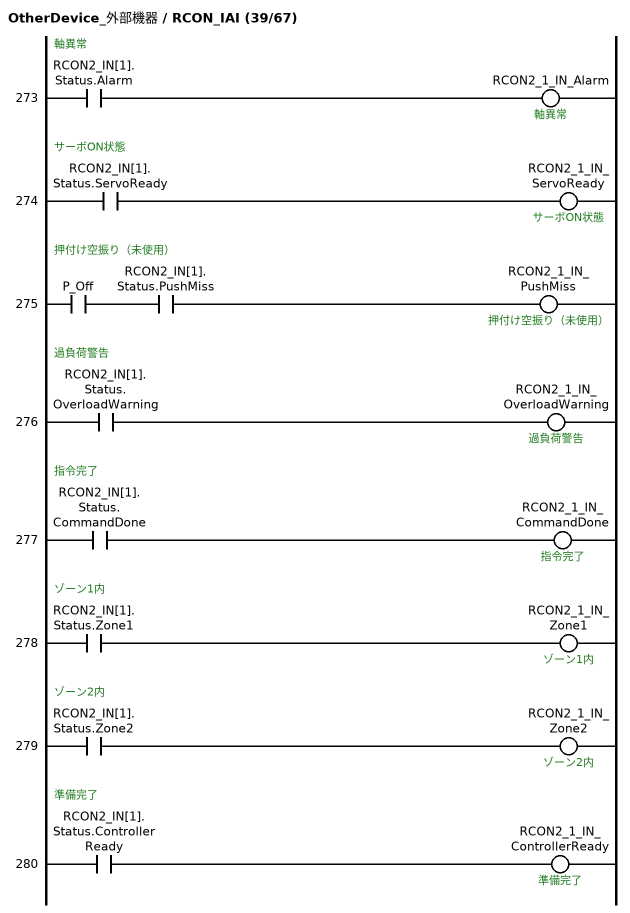
(* Rung 273: 軸異常 *)
RCON2_1_IN_Alarm := RCON2_IN[1].Status.Alarm;
(* Rung 274: サーボON状態 *)
RCON2_1_IN_ServoReady := RCON2_IN[1].Status.ServoReady;
(* Rung 275: 押付け空振り（未使用） *)
RCON2_1_IN_PushMiss := P_Off AND RCON2_IN[1].Status.PushMiss;
(* Rung 276: 過負荷警告 *)
RCON2_1_IN_OverloadWarning := RCON2_IN[1].Status.OverloadWarning;
(* Rung 277: 指令完了 *)
RCON2_1_IN_CommandDone := RCON2_IN[1].Status.CommandDone;
(* Rung 278: ゾーン1内 *)
RCON2_1_IN_Zone1 := RCON2_IN[1].Status.Zone1;
(* Rung 279: ゾーン2内 *)
RCON2_1_IN_Zone2 := RCON2_IN[1].Status.Zone2;
(* Rung 280: 準備完了 *)
RCON2_1_IN_ControllerReady := RCON2_IN[1].Status.ControllerReady;

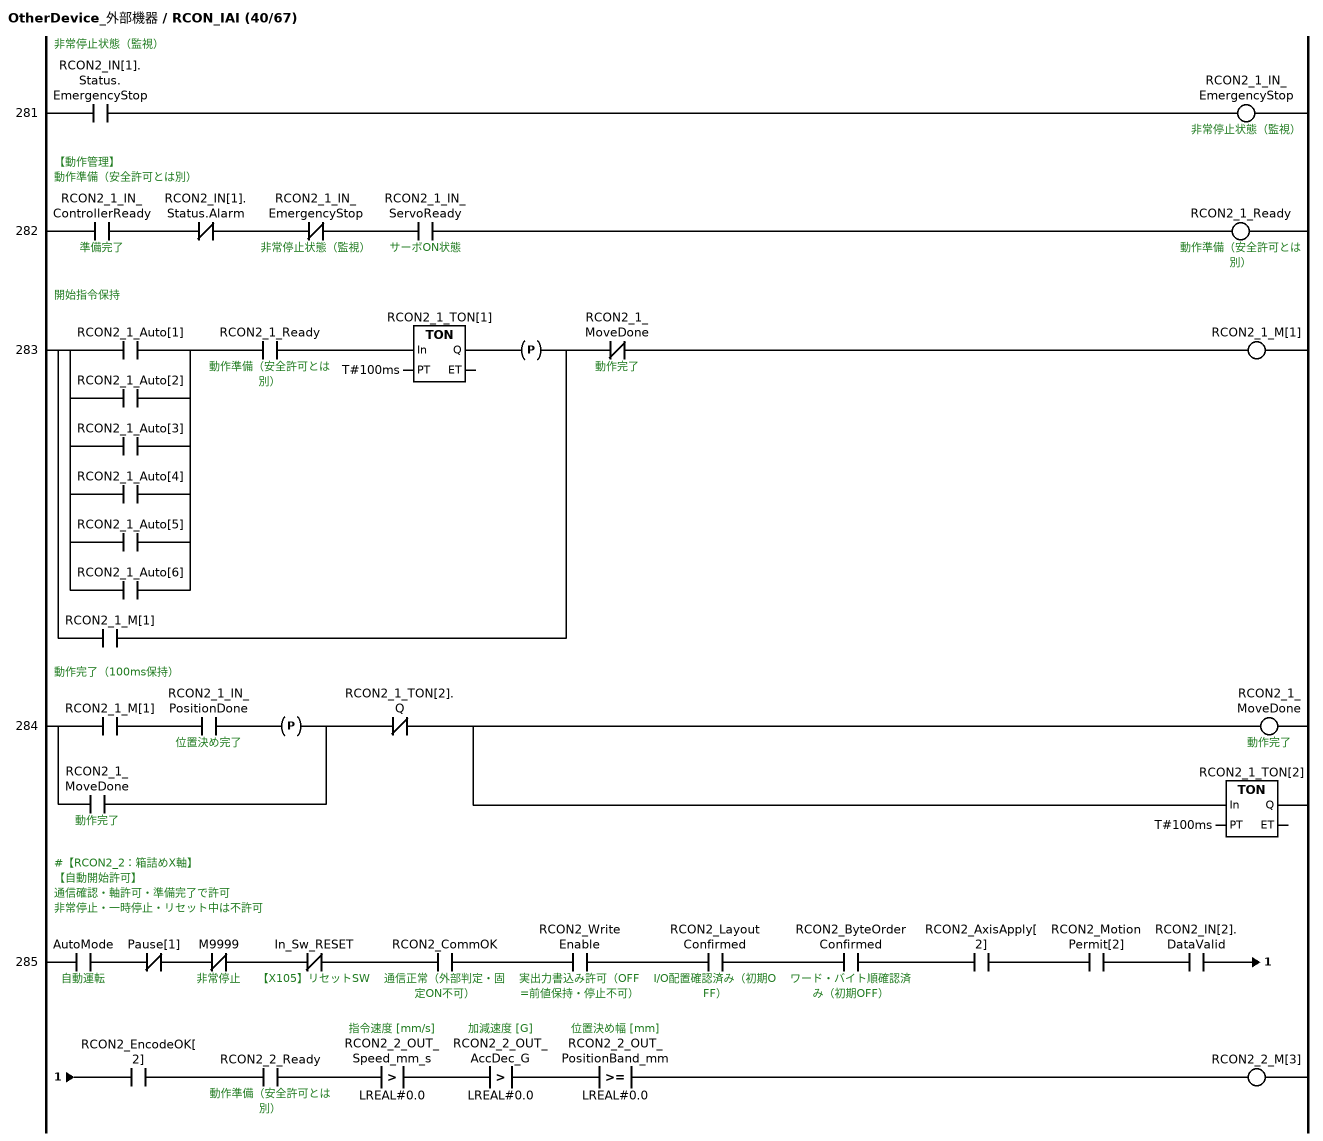
(* Rung 281: 非常停止状態（監視） *)
RCON2_1_IN_EmergencyStop := RCON2_IN[1].Status.EmergencyStop;
(* Rung 282: 【動作管理】 / 動作準備（安全許可とは別） *)
RCON2_1_Ready := RCON2_1_IN_ControllerReady AND NOT RCON2_IN[1].Status.Alarm AND NOT RCON2_1_IN_EmergencyStop AND RCON2_1_IN_ServoReady;
(* Rung 283: 開始指令保持 *)
RCON2_1_TON[1](In := (RCON2_1_Auto[1] OR RCON2_1_Auto[2] OR RCON2_1_Auto[3] OR RCON2_1_Auto[4] OR RCON2_1_Auto[5] OR RCON2_1_Auto[6]) AND RCON2_1_Ready, PT := T#100ms);
_e26(CLK := RCON2_1_TON[1].Q);
RCON2_1_M[1] := (_e26.Q OR RCON2_1_M[1]) AND NOT RCON2_1_MoveDone;
(* Rung 284: 動作完了（100ms保持） *)
_e27(CLK := RCON2_1_M[1] AND RCON2_1_IN_PositionDone);
_p28 := (_e27.Q OR RCON2_1_MoveDone) AND NOT RCON2_1_TON[2].Q;
RCON2_1_MoveDone := _p28;
RCON2_1_TON[2](In := _p28, PT := T#100ms);
(* Rung 285: #【RCON2_2：箱詰めX軸】 / 【自動開始許可】 / 通信確認・軸許可・準備完了で許可 / 非常停止・一時停止・リセット中は不許可 *)
RCON2_2_M[3] := AutoMode AND NOT Pause[1] AND NOT M9999 AND NOT In_Sw_RESET AND RCON2_CommOK AND RCON2_WriteEnable AND RCON2_LayoutConfirmed AND RCON2_ByteOrderConfirmed AND RCON2_AxisApply[2] AND RCON2_MotionPermit[2] AND RCON2_IN[2].DataValid AND RCON2_EncodeOK[2] AND RCON2_2_Ready AND (RCON2_2_OUT_Speed_mm_s > LREAL#0.0) AND (RCON2_2_OUT_AccDec_G > LREAL#0.0) AND (RCON2_2_OUT_PositionBand_mm >= LREAL#0.0);

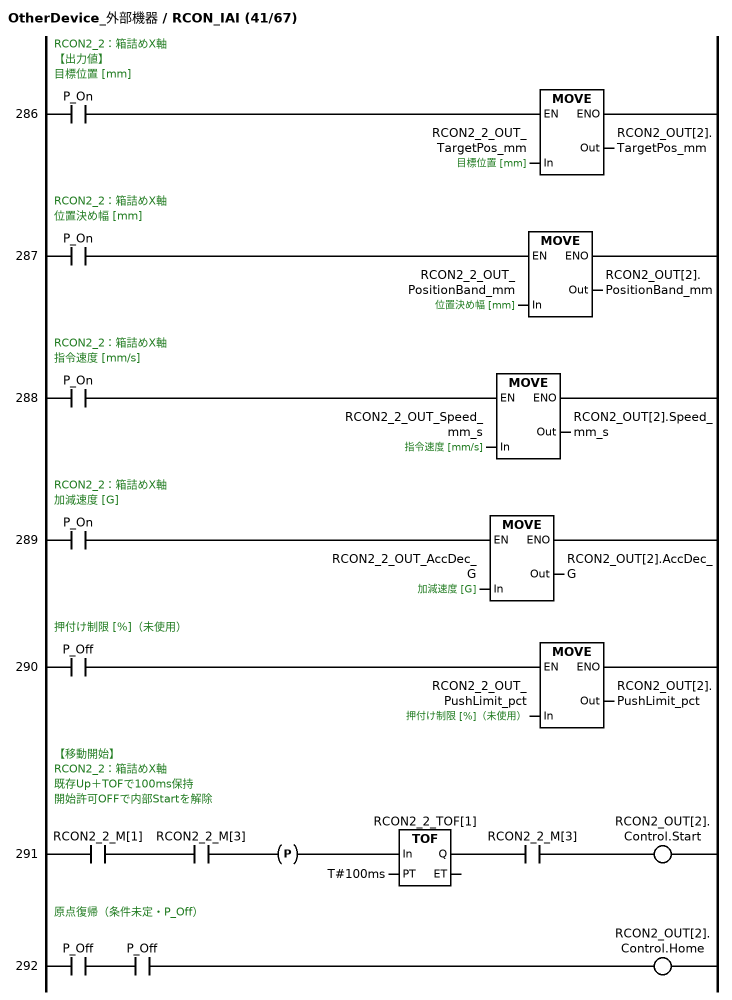
(* Rung 286: RCON2_2：箱詰めX軸 / 【出力値】 / 目標位置 [mm] *)
IF P_On THEN RCON2_OUT[2].TargetPos_mm := RCON2_2_OUT_TargetPos_mm; END_IF;
(* Rung 287: RCON2_2：箱詰めX軸 / 位置決め幅 [mm] *)
IF P_On THEN RCON2_OUT[2].PositionBand_mm := RCON2_2_OUT_PositionBand_mm; END_IF;
(* Rung 288: RCON2_2：箱詰めX軸 / 指令速度 [mm/s] *)
IF P_On THEN RCON2_OUT[2].Speed_mm_s := RCON2_2_OUT_Speed_mm_s; END_IF;
(* Rung 289: RCON2_2：箱詰めX軸 / 加減速度 [G] *)
IF P_On THEN RCON2_OUT[2].AccDec_G := RCON2_2_OUT_AccDec_G; END_IF;
(* Rung 290: 押付け制限 [%]（未使用） *)
IF P_Off THEN RCON2_OUT[2].PushLimit_pct := RCON2_2_OUT_PushLimit_pct; END_IF;
(* Rung 291: 【移動開始】 / RCON2_2：箱詰めX軸 / 既存Up＋TOFで100ms保持 / 開始許可OFFで内部Startを解除 *)
_e29(CLK := RCON2_2_M[1] AND RCON2_2_M[3]);
RCON2_2_TOF[1](In := _e29.Q, PT := T#100ms);
RCON2_OUT[2].Control.Start := RCON2_2_TOF[1].Q AND RCON2_2_M[3];
(* Rung 292: 原点復帰（条件未定・P_Off） *)
RCON2_OUT[2].Control.Home := P_Off AND P_Off;

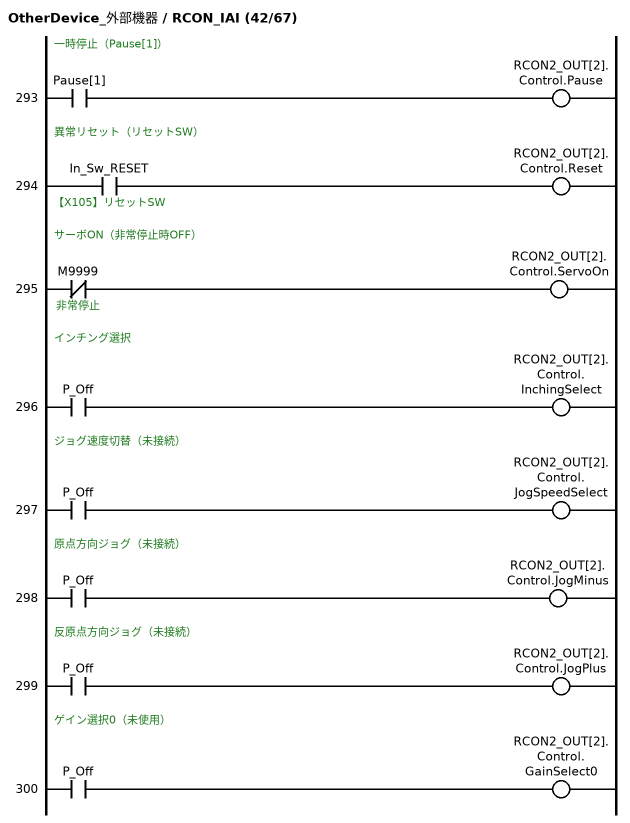
(* Rung 293: 一時停止（Pause[1]） *)
RCON2_OUT[2].Control.Pause := Pause[1];
(* Rung 294: 異常リセット（リセットSW） *)
RCON2_OUT[2].Control.Reset := In_Sw_RESET;
(* Rung 295: サーボON（非常停止時OFF） *)
RCON2_OUT[2].Control.ServoOn := NOT M9999;
(* Rung 296: インチング選択 *)
RCON2_OUT[2].Control.InchingSelect := P_Off;
(* Rung 297: ジョグ速度切替（未接続） *)
RCON2_OUT[2].Control.JogSpeedSelect := P_Off;
(* Rung 298: 原点方向ジョグ（未接続） *)
RCON2_OUT[2].Control.JogMinus := P_Off;
(* Rung 299: 反原点方向ジョグ（未接続） *)
RCON2_OUT[2].Control.JogPlus := P_Off;
(* Rung 300: ゲイン選択0（未使用） *)
RCON2_OUT[2].Control.GainSelect0 := P_Off;

